Fanuc KAREL source: KA00168.KL

PROGRAM KA00168
%NOLOCKGROUP
VAR
  SRC: ARRAY[4] OF BOOLEAN
  DST: ARRAY[4] OF SHORT
BEGIN
  DST = SRC
END KA00168
